Fanuc KAREL source: KA00157.KL

PROGRAM KA00157
%NOLOCKGROUP
VAR
  SRC: ARRAY[4] OF REAL
  DST: ARRAY[4] OF STRING[20]
BEGIN
  DST = SRC
END KA00157
